(* IEC 61131-3 sources: plc-vscode/tests/st/all/trust-platform/manual-tests/root-b/src, 1 file *)

(* ---- Other.st ---- *)
PROGRAM Main
VAR
    value : DINT;
END_VAR
value := 42;
END_PROGRAM
